Fanuc KAREL source: ke00004.KL

-- PROVISIONAL review KL for V1013-1; original PC SHA256 ca5c5950b72b9f582d9b294dadbcb4a6dbbe206b688bbe85a1b2e9bac58c870f
-- Incomplete behavior may be omitted. Consult companion uncertainty JSON. Do not deploy.
PROGRAM KE00004
%NOLOCKGROUP
BEGIN
  -- UNRESOLVED_PC offsets 5-12; opcodes 9D,23
  -- UNRESOLVED_PC offsets 17-29; opcodes 3F,75
  -- UNRESOLVED_PC offsets 34-58; opcodes 27,22,22,2A,22,31
  -- UNRESOLVED_PC offsets 63-67; opcodes 7F
END KE00004
